(* IEC 61131-3 sources: Versio-VersionControlSystem/fixtures/projects/TC3_PlcSample_reStrText/TC3_PlcSample_reStrText/LibraryDocumentationSample Project/LibPOUs/B_DocuElements/Font style, 1 file *)

(* ---- FB_Libdoc_FontStyle.st ---- *)
(*
This is *emphasized text*.

This is **strong text**.

This text is an example of ``inline literals``.
*)

FUNCTION_BLOCK FB_Libdoc_FontStyle
VAR_INPUT
    nVarA : INT;
    nVarB : INT;
END_VAR
VAR_OUTPUT
    nSum : INT;
END_VAR
VAR
END_VAR
